// LS Electric XG5000 project: cell
// PLC LSPLC

PROGRAM NewProgram (task: Scan Program)

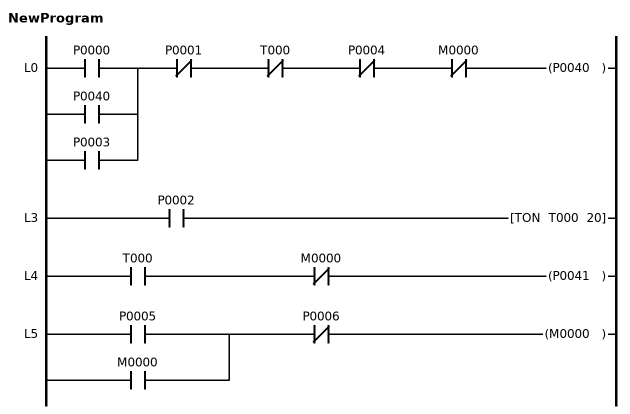
; L0
LOAD      P0000
OR        P0040
OR        P0003
AND NOT   P0001
AND NOT   T000
AND NOT   P0004
AND NOT   M0000
OUT       P0040
; L3
LOAD      P0002
TON       T000 20
; L4
LOAD      T000
AND NOT   M0000
OUT       P0041
; L5
LOAD      P0005
OR        M0000
AND NOT   P0006
OUT       M0000